TYPE ST_VisuFingerState :
STRUCT
	stPose : ST_VisuPose; // MCS, absolute: pose of the finger's frame (centre of its top face)
	(* The application reported stPose (protocol 20, ADR 0018). FALSE: clients place the finger by its stOffset on
	   the gripper flange. Set by the library, not by the application. *)
	bPoseReported : BOOL;
	bActive : BOOL; // the finger grips
END_STRUCT
END_TYPE

(* stored: Version 1.1.0.1, ProductVersion 3.1.4026.18
   DUT ST_VisuFingerState: Id {8b376170-d812-4be6-8c74-d7d224b9dfd4} *)
